// TIA Portal V19 export
TYPE "FctKeyParName"
   STRUCT
      Key : UInt;
      "Name" : String;
   END_STRUCT;
END_TYPE
